(* IEC 61131-3 sources: Caravan/Archiv/12-04-19/Stations/MachineControl/MachineControl/Class/LseEasy (part 2) *)

  if(input < 0) then
    input := 0;
    result := ACCESS_DENIED;
  elsif(input > 100) then
    input := 100;
    result := ACCESS_DENIED;
  else
	  result := input;
  end_if;

  ComPort.SendBacklightDim(input$usint);
	BacklightDim := input;

END_FUNCTION

FUNCTION LseEasy::GetBacklightDim
	VAR_OUTPUT
		retcode 	: USINT;
	END_VAR

  retcode := ComPort.GetBacklightInfo();
  if(retcode <> 0xFF) then
    BacklightDim := retcode and 0x7F;
  end_if;

END_FUNCTION

FUNCTION GLOBAL LseEasy::UpdateScreenshot
	VAR_INPUT
		pscrshot 	: ^void;
	END_VAR

  if(ComPort.SaveScreenshot("C:\hmi35.bmp", pscrshot) = true) then
    OutMessage("SCREENSHOT ...Ready (C:\hmi35.bmp)");
  else
    OutMessage("ERROR: Can't save Screenshot (C:\hmi35.bmp)");
  end_if;

  if(StateSvr = TGetScreenShot) then
    StateSvr := TRun;
  end_if;

END_FUNCTION

FUNCTION VIRTUAL GLOBAL LseEasy::UpdateValue35
	VAR_INPUT
		varno 	: UINT;
		value 	: DINT;
	END_VAR

  if(HmiPrjCrc = Hmi35PrjCrc) then // check crc of project with crc of hmi

    if(varno = VARNO_IRCODE) then
      UpdateIrCode(value$udint);
    end_if;

    HmiVarList.UpdateValue(varno, value);
  end_if;

END_FUNCTION

FUNCTION VIRTUAL GLOBAL LseEasy::UpdateString35
	VAR_INPUT
		varno 	: UINT;
		pstr 	: ^void;
		chrsize 	: UDINT;
	END_VAR

  if(HmiPrjCrc = Hmi35PrjCrc) then // check crc of project with crc of hmi
    HmiVarList.UpdateString(varno, pstr, chrsize);
  end_if;

END_FUNCTION

FUNCTION VIRTUAL GLOBAL LseEasy::UpdateTemperature35
	VAR_INPUT
		value 	: DINT;
	END_VAR

  ActTemperature := value;

END_FUNCTION

FUNCTION GLOBAL LseEasy::UpdateActScreen
	VAR_INPUT
		scrno 	: DINT;
	END_VAR

  ActScreen := scrno;

END_FUNCTION

FUNCTION GLOBAL LseEasy::UpdateInUse

  LastUsage := ops.tAbsolute;

END_FUNCTION

FUNCTION VIRTUAL GLOBAL LseEasy::ActLanguage::Write
	VAR_INPUT
		input (EAX) 	: UDINT;
	END_VAR
	VAR_OUTPUT
		result (EAX) 	: UDINT;
	END_VAR

  if(input <> ActLanguage) then
    if(HmiTextList.GetLanguageIndex(input) <> 16#FFFFFFFF) then
	    ActLanguage := input;
      if(StateSvr = TRun) then
        StateSvr := TStart;
      end_if;
    end_if;
  end_if;

	result := ActLanguage;

END_FUNCTION

FUNCTION GLOBAL LseEasy::SendNewBootLoader
	VAR_OUTPUT
		retcode 	: bool;
	END_VAR

  retcode := SendUpdateToHmi(GetBootLoaderUpdate());

END_FUNCTION

FUNCTION GLOBAL LseEasy::SendNewFirmware
	VAR_OUTPUT
		retcode 	: bool;
	END_VAR

  retcode := SendUpdateToHmi(GetFirmwareUpdate());

END_FUNCTION

FUNCTION LseEasy::SendUpdateToHmi
	VAR_INPUT
		dpne 	: ^CHAR;
	END_VAR
	VAR_OUTPUT
		retcode 	: BOOL;
	END_VAR
  VAR
  	length : udint;
    pbin : ^void;
    tmp : array[0..300] of char;
  END_VAR

  retcode := false;
  pbin    := NIL;

  ComPort.SendBacklightOnOff(1); // turn on backlight

  StringLib.StrCpy(#tmp, 1, "FIRMWARE-UPDATE: Start...[", 1);
  StringLib.StrCat(#tmp, 1, dpne, 1);
  StringLib.StrCat(#tmp, 1, "]", 1);
  OutMessage(#tmp[0]);

  if(File.FOpen(dpne, 'r') = true) then
    length$dint := File.FLength();
    if(length$dint > 0) then
      if(File.FMemory(#pbin, length + 4) = true) then
        if(File.FRead(pbin+4, length) = true) then
          pbin$^udint^ := CRC32_Buffer(pbin+4, length);
          retcode := ComPort.SendNewFirmware(pbin, length+4);
          if(retcode = false) then
            StringLib.StrCpy(#tmp[0], sizeof(char), "ERROR: can't upload ", sizeof(char));
            StringLib.StrCat(#tmp[0], sizeof(char), dpne, sizeof(char));
            OutMessage(#tmp[0]);
          end_if;
        end_if;
        File.FMemory(#pbin, 0);
      end_if;
    end_if;
  else
    StringLib.StrCpy(#tmp[0], sizeof(char), "ERROR: can't open ", sizeof(char));
    StringLib.StrCat(#tmp[0], sizeof(char), dpne, sizeof(char));
    OutMessage(#tmp[0]);
  end_if;

  File.FClose();

  if(retcode = true) then
    OutMessage("FIRMWARE-UPDATE: ...Ready");
  end_if;

END_FUNCTION

FUNCTION GLOBAL LseEasy::SendTrend
	VAR_INPUT
		id 	: UDINT;
		pdata 	: ^USINT;
		length 	: UDINT;
	END_VAR

  ComPort.SendTrendValue(id, pdata, length);

END_FUNCTION

FUNCTION GLOBAL LseEasy::SendPixMap
	VAR_INPUT
		pdata 	: ^void;
		width 	: USINT;
		height 	: USINT;
		padding 	: USINT;
	END_VAR
	VAR_OUTPUT
		retcode 	: BOOL;
	END_VAR
  VAR
  	size : udint;
  END_VAR

  retcode := false;
  size    := ((width * height) + 7) / 8;
  size    += 5; // headerdaten

  // [] ..... command
  // [] ..... version = 1
  // [] ..... width
  // [] ..... height
  // [] ..... padding
  // [ ...... bitdata

  if(size <= sizeof(TmpData)) then
    TmpData[0] := ComCMD_UPDATEPIXMAP;
    TmpData[1] := 1;
    TmpData[2] := width;
    TmpData[3] := height;
    TmpData[4] := padding;
    MemCpy3(#TmpData[5], pdata, size-5);
    retcode := ComPort.SendData(#TmpData[0], size);
  end_if;

END_FUNCTION

FUNCTION GLOBAL LseEasy::OutMessage
	VAR_INPUT
		txt 	: ^CHAR;
	END_VAR
  VAR
  	tmp : array[0..300] of char;
  END_VAR

  tmp[0] := '[';
  tmp[1] := 'N';
  tmp[2] := 'o';
  tmp[3] := 'd';
  tmp[4] := 'e';
  tmp[5] := ' ';
  StringLib.DintToStr(#tmp[6], to_int(ComPort.GetNode()), 16#0800, 1);
  StringLib.StrCat(#tmp[6], 1, "] ", 1);
  StringLib.StrCat(#tmp[6], 1, txt, 1);
  TRACE(#tmp[0]);

END_FUNCTION

FUNCTION LseEasy::OutMessageValue
	VAR_INPUT
		txt 	: ^CHAR;
    value : udint;
	END_VAR
  VAR
  	msg : array[0..128] of char;
  END_VAR

  StringLib.StrCpy(#msg[0], 1, txt, 1);
  StringLib.DintToStr(#msg[StringLib.StrLen(#msg[0], 1)], to_dint(value), 0x800, 1);
  OutMessage(#msg[0]);

END_FUNCTION

FUNCTION GLOBAL LseEasy::UpdateAll
	VAR_INPUT
		act_hmi_crc 	: UDINT;
	END_VAR

  Hmi35PrjCrc   := act_hmi_crc;
  NeedUpdateAll += 1;

END_FUNCTION

FUNCTION LseEasy::CheckCrc
VAR
	crc : udint;
END_VAR

  crc := ComPort.GetFileCrc(0);
  if(crc = 16#FFFFFFFF) then
    // there is no valid project in hmi
    StateSvr := TStart; // restart
  elsif(crc <> 0) then
    CantGetCrc := 0;
    if(crc = HmiPrjCrc) then
      // same project detected in hmi
      UpdateAll(crc); // force update of all data
      StateSvr := TRun;
    else
      // different project detected in hmi
      StateSvr := TStart; // restart
    end_if;
  else

    SleepNext(StateSvr, 100); // sleep 100ms

    CantGetCrc += 1;
    if(CantGetCrc > 100) then
      CantGetCrc := 0;
      ErrorStateSvr(true);
    end_if;
  end_if;

END_FUNCTION

FUNCTION GLOBAL LseEasy::UpdateAliveSignal35

  AliveTix35     := ops.tAbsolute;
  HmiOnline      := 1;
  AliveTix35Cntr += 1;

END_FUNCTION

FUNCTION GLOBAL LseEasy::UpdateBacklight35
	VAR_INPUT
		state 	: DINT;
	END_VAR

//  if(state and 0x80) then
//    BacklightOnOff := 1;
//  else
//    BacklightOnOff := 0;
//  end_if;

  BacklightDim := state and 0x7F;

END_FUNCTION

FUNCTION LseEasy::CheckProjectCrc
	VAR_INPUT
		ptr 	: ^void;
		hmiver 	: UDINT;
		chkold 	: bool;
	END_VAR
	VAR_OUTPUT
		retcode 	: BOOL;
	END_VAR
  VAR
  	pprj : ^_BOX_PROJECTLIST;
  	phlp : ^_BOX_PROJECTLIST_ENTRY;
    no, index : udint;
		pbox	: ^_BIGBOX_HEADER;
    upload : bool;
  END_VAR

  upload     := true;
  retcode    := false;
  pbox$^void := ptr;

  if(ComPort.GetFileCrc(0) = pbox^.crc32) then
    retcode := true;
    upload  := false;
    if((chkold = true) & (hmiver < 127)) then
      // einzelne crc's im hmi überprüfen
      // erst ab hmi-version 1.27 werden die crc's mit GetFileCrc(0) direkt im hmi überprüft
      pprj$^void := pbox;
      no         := pprj^.no;
      phlp       := #pprj^.data[0];
      index      := 0;

      while(no) do
        no    -= 1;
        pbox$^void := HmiProject35.GetBox(index);

        if(ComPort.GetFileCrc(phlp^.filename) <> pbox^.crc32) then
          retcode := false;
          no      := 0;
        end_if;

        phlp  += sizeof(_BOX_PROJECTLIST_ENTRY);
        index += 1;
      end_while;
    end_if;
  end_if;

  if(IsProjectUpLoadNecessary(upload) = true) then
    retcode := false;
  end_if;

END_FUNCTION

FUNCTION LseEasy::SendProject
	VAR_INPUT
		ptr 	: ^void;
	END_VAR
	VAR_OUTPUT
		retcode 	: BOOL;
	END_VAR
  VAR
  	pprj : ^_BOX_PROJECTLIST;
  	phlp : ^_BOX_PROJECTLIST_ENTRY;
    no, index, tix, nox, sizeram, sizeflash : udint;
    pbox : ^_BIGBOX_HEADER;
    upload : bool;
  END_VAR

  retcode := false;
  upload  := false;

  tix := ops.tAbsolute;

    if(ComPort.SendReset() = true) then

      HmiSwVersion := ComPort.GetSwVersion();
      HmiHwVersion := ComPort.GetHwVersion();

      GetBacklightDim();

      pbox$^void := ptr;
      retcode    := true;

      // nur wenn projektcrc unterschiedlich
      if(CheckProjectCrc(ptr, HmiSwVersion, false) = false) then

        if(ComPort.GetHardwareData(nil, #sizeram, #sizeflash) = true) then
          sizeflash := sizeflash - (24 + 512*16); // flashhader + fatgrösse abziehen
          if((HmiProject35.TotalByteSize > sizeflash) | (HmiProject35.TotalFileNo > 256)) then
            OutMessage("ERROR: Size of LSE-Project is too big");
            OutMessageValue("...PrjSize[byte] = ", HmiProject35.TotalByteSize);
            OutMessageValue("...MaxSize[byte] = ", sizeflash);
            SetErrorSvr(ErrSizeLseProject);
            retcode := false;
          end_if;
        end_if;

        if(retcode = true) then

          // clear flash
          if(ComPort.SendFormatFlash() = true) then

            OutMessage("HMI-UPDATE: Start...");

            // send projectentries
            pprj$^void := ptr;
            no         := pprj^.no;
            phlp       := #pprj^.data[0];
            index      := 0;
//            totalsize  := 0;

            while(no) do
              ComPort.ShowProgressBar(to_usint((index * 100) / pprj^.no));

              no    -= 1;
              pbox$^void := HmiProject35.GetBox(index);

              if(ComPort.SendFile(phlp^.filename, pbox^.size, pbox) = false) then
                OutMessageValue("ERROR: Upload ProjectEntry of Bytesize = ", pbox^.size);
                retcode := false;
                no      := 0;
              end_if;
//              totalsize += HmiProject35.AlignU32(pbox^.size);
              phlp  += sizeof(_BOX_PROJECTLIST_ENTRY);
              index += 1;
            end_while;

            if(retcode = true) then
              // send projektlist
              ComPort.ShowProgressBar(100);
              pbox$^void := ptr;
              retcode    := ComPort.SendFile(0, pbox^.size, pbox);
//              totalsize  += HmiProject35.AlignU32(pbox^.size);

              if(retcode = true) then
                HmiMapFile.Create(GetPrjPath(), pbox^.crc32);
                OutMessageValue("HMI-UPDATE: ...Ready, TotalSize[byte] = ", HmiProject35.TotalByteSize); //totalsize);
                // vorsicht: projekt ist jetzt im hmi-ram, noch nicht auf flash
                retcode := ComPort.Ping(); // send ping to ensure alive-hmi and update alivetrigger
              end_if;
              upload := true;
            end_if;

          else
            retcode := false;
          end_if;
        end_if;
      end_if;

      if(retcode = true) then
        UpdateAll(HmiPrjCrc); // force updateall
        nox := ops.tAbsolute;
        repeat
          if(ComPort.SendRun() = true) then
            exit;
          end_if;
        until((ops.tAbsolute - nox) > 1000) end_repeat;

        if(upload = true) then
          // after performing projectupload, sleep a while to ensure flash of whole project-data in hmi
          nox := ops.tAbsolute;
          while((ops.tAbsolute - nox) < 1000) do
          end_while;
          ComPort.Ping(); // send ping to keep hmi happy
        end_if;

        OutMessageValue("HMI-RUN: UpdateTime[ms] = ", ops.tAbsolute - tix);
      else
        OutMessage("ERROR: Upload HMI-Project");
        SetErrorSvr(ErrUploadHmiProject);
        ComPort.SendChkTraceView(); // display message on hmi
      end_if;
    end_if;

END_FUNCTION

FUNCTION LseEasy::Run

  // alivesignal
  if((ops.tabsolute - AliveTix) > 1003) then
    AliveTix := ops.tabsolute;
    ComPort.SendAliveTrigger(); // send alive trigger to hmi
  end_if;

  // onlinewatchdog
  if((ops.tabsolute - AliveTix35) > 4000) then
    HmiOnline := 0; // offline
    if(TempInterval <> 0) then
      ActTemperature$UDINT := 0x80000010; // fühlerbruch
    end_if;
  end_if;

  if(HmiOnline) then

    if(HmiPrjCrc = Hmi35PrjCrc) then // check crc of project with crc of hmi

      if(NeedUpdateAll) then
        NeedUpdateAll := 0;
        GetBacklightDim();
        HmiVarList.RefreshAll();
        HmiStateBit35.RefreshAll();
        HmiReady();
      end_if;

      HmiRun();

      if((ops.tabsolute - RefreshTix) > 6) then
        RefreshTix := ops.tAbsolute;
        HmiVarList.RefreshRun();
        HmiStateBit35.RefreshRun();
      end_if;

      if(TrendVal0 <> -1) then
        TrendVal0 := UpdateTrendVal(0, TrendVal0);
      end_if;

      if(TrendVal1 <> -1) then
        TrendVal1 := UpdateTrendVal(1, TrendVal1);
      end_if;

      if(PixMap <> -1) then
        PixMap := UpdatePixMap(PixMap);
      end_if;

    else
      // just in this moment we're back online with hmi
      SleepNext(TChkCrc, 1000); // wait a while and afterwards check project
    end_if;
  else
    Hmi35PrjCrc := 0; // destroy hmicrc
    CantGetCrc  := 0;
  end_if;

  if(CallScreen <> -1) then
    if(CallScreen = -2) then
      OutMessage("SCREENSHOT: Start...");
      if(ComPort.GetScreenShot() = false) then
        OutMessage("ERROR: Screenshot not done");
      else
        StateSvr := TGetScreenShot;
      end_if;
    else
      ComPort.SendGotoScreen(CallScreen);
    end_if;
    CallScreen := -1;
  end_if;

END_FUNCTION

FUNCTION VIRTUAL GLOBAL LseEasy::Background
	VAR_INPUT
		EAX 	: UDINT;
	END_VAR
	VAR_OUTPUT
		state (EAX) 	: UDINT;
	END_VAR

	state := READY;

  case StateSvr of
    TStart :
      AutoFirmwareUpdate := AutoFirmwareUpdate.Read();
      if(ComPort.Ping() = true) then // ask for hmi
        if(LoadFile() = true) then
          if(Create() = true) then
            StateSvr := TUpload;
          end_if;
        end_if;

        if(StateSvr <> TUpload) then
          ErrorStateSvr(false);
        else
          if(AutoFirmwareUpdate <> 0) then
            if(AutoFwUpdateDisabled = false) then
              AutoFwUpdateDisabled := true; // no further auto-update of firmware possible
              StateSvr := TCheckUpdateBootloader;
            end_if;
          end_if;
        end_if;
      else
        OutMessage("ERROR: Can't communicate with HMI");
        SetErrorSvr(ErrHmiCommunication);
        ErrorStateSvr(true);
      end_if;

    TCheckUpdateBootLoader :
      StateSvr := CheckUpdate(GetBootloaderUpdate(), TCheckUpdateFirmware, TCheckUpdateFirmware, 15000);

    TCheckUpdateFirmware :
      StateSvr := CheckUpdate(GetFirmwareUpdate(), TStart, TUpLoad, 17000);

    TUpLoad :
      if(UpLoadProject() = true) then
        HmiProject35.Free();
        ProjectBox := NIL;
        StateSvr := TRun;
      end_if;

    TGetScreenShot :
      Run();

    TRun :
      Run();

    TFirmwareUpdate :
      if(SendNewFirmware() = true) then
        SleepNext(TRun, 10000);
      else
        ErrorStateSvr(false);
      end_if;

    TBootLoaderUpdate :
      if(SendNewBootLoader() = true) then
        SleepNext(TRun, 10000);
      else
        ErrorStateSvr(false);
      end_if;

    TChkCrc :
      CheckCrc();

    TSleep :
      if((ops.tAbsolute - SleepStart) >= SleepDuration) then
        StateSvr := StateNext;
      end_if;

    TReboot :
      ComPort.SendReboot();
      SleepNext(TStart, 3000);

    TError :
      if(TryToRestart = true) then
        if(AliveTix35Cntr <> AliveTix35CntrOld) then
          // try to restart after hmi sent alivesignal
          StateSvr     := TStart;
          TryToRestart := false;
        end_if;
      end_if;

  end_case;

  ComPort.Run();

END_FUNCTION

FUNCTION VIRTUAL GLOBAL LseEasy::StateSvr::Write
	VAR_INPUT
		input (EAX) 	: LseEasy::TStateSvr;
	END_VAR
	VAR_OUTPUT
		result (EAX) 	: LseEasy::TStateSvr;
	END_VAR

  if(input = TGetScreenShot) then
    result$udint := ACCESS_DENIED;
    if(StateSvr = TRun) then
      CallScreen := -2;
	    result     := StateSvr;
    end_if;
  else
	  StateSvr := input;
	  result := StateSvr;
  end_if;

END_FUNCTION

FUNCTION VIRTUAL GLOBAL LseEasy::HmiAccess
	VAR_INPUT
		level 	: UDINT;
	END_VAR
	VAR_OUTPUT
		retcode 	: BOOL;
	END_VAR

  retcode := true;
  if(level > AccessLevel) then
    retcode := false;
  end_if;

END_FUNCTION

FUNCTION GLOBAL LseEasy::SoftReset

  StateSvr := TStart;

END_FUNCTION

FUNCTION GLOBAL LseEasy::SoftResetAll
  VAR
  	nox : udint;
    pth : ^LseEasy;
  END_VAR

  pth := InstancePtr[0];
  nox := InstanceCnt;
  while(nox) do
    pth^.SoftReset();
    nox -= 1;
    pth += sizeof(InstancePtr[0]);
  end_while;

END_FUNCTION

FUNCTION VIRTUAL GLOBAL LseEasy::ClassSvr::NewInst
	VAR_INPUT
		pPara 	: ^CmdStruct;
		pResult 	: ^Results;
	END_VAR
	VAR_OUTPUT
		ret_code 	: IprStates;
	END_VAR

	ret_code := READY;

	case pPara^.uiCmd of

		0 : // start download on the fly
        pResult^.aData[0]$UDINT := 16#46544F44; // DOTF-id
        pResult^.uiLng          := 6; // success

		1 : // end download on the fly
        pResult^.aData[0]$UDINT := 16#46544F44; // DOTF-id
        pResult^.uiLng          := 6; // success
        SoftResetAll();
  end_case;

END_FUNCTION

#pragma warning (disable : 73)
FUNCTION VIRTUAL GLOBAL LseEasy::UserCall
	VAR_INPUT
		fktno 	: UDINT;
		para 	: DINT;
	END_VAR

END_FUNCTION
#pragma warning (default : 73)

#pragma warning (disable : 73)
FUNCTION VIRTUAL GLOBAL LseEasy::HmiVariableExtention
	VAR_INPUT
		varname 	: ^CHAR;
	END_VAR
	VAR_OUTPUT
		retcode 	: UDINT;
	END_VAR

  retcode := 16#FFFFFFFF;

//  if(StringLib.StrCmp(varname, sizeof(char), "Dummy.Server7", sizeof(char)) = 0) then
//    retcode := VARNO_TEST_NUM1;
//  end_if;

END_FUNCTION
#pragma warning (default : 73)

FUNCTION LseEasy::GetMapCrc
	VAR_OUTPUT
		retcode 	: UDINT;
	END_VAR

  retcode := HmiVarList.GetMapCrc();
  retcode := (retcode rol 1) xor HmiStateBit35.GetMapCrc();

END_FUNCTION

FUNCTION VIRTUAL LseEasy::IsProjectUpLoadNecessary
	VAR_INPUT
		preselect 	: BOOL;
	END_VAR
	VAR_OUTPUT
		retcode 	: BOOL;
	END_VAR

//  if(GetmapCrc() <> oldmapcrc) then
    // unconditional upload necessary, otherwise weak functionality of hmi
//  end_if;

  retcode := preselect;

END_FUNCTION

FUNCTION VIRTUAL GLOBAL LseEasy::UpdatePixMap
	VAR_INPUT
		value 	: DINT;
	END_VAR
	VAR_OUTPUT
		retcode 	: DINT;
	END_VAR

  retcode := value;
  if(SendPixMap(#value, 32, 1, 0) = true) then
    retcode := -1;
  end_if;

END_FUNCTION

FUNCTION VIRTUAL GLOBAL LseEasy::UpdateTrendVal
	VAR_INPUT
    id : UDINT;
		value 	: DINT;
	END_VAR
	VAR_OUTPUT
		retcode 	: DINT;
	END_VAR

  retcode := value;
  if(ComPort.SendTrendValue(id, #(value$usint), 1) = true) then
    retcode := -1;
  end_if;

END_FUNCTION

FUNCTION LseEasy::Recalculate_MulDiv
	VAR_INPUT
		einheit 	: UDINT;
		posdezpt 	: DINT;
	END_VAR
	VAR_OUTPUT
		retcode 	: DINT;
	END_VAR
  var
    dekade : dint;
  end_var

  retcode := 1;
  dekade  := 0;

  case(einheit) of
    1000000000 : dekade := 9;
    100000000  : dekade := 8;
    10000000   : dekade := 7;
    1000000    : dekade := 6;
    100000     : dekade := 5;
    10000      : dekade := 4;
    1000       : dekade := 3;
    100        : dekade := 2;
    10         : dekade := 1;
  end_case;

  case(dekade - posdezpt) of
    9 : retcode := 1000000000;
    8 : retcode :=  100000000;
    7 : retcode :=   10000000;
    6 : retcode :=    1000000;
    5 : retcode :=     100000;
    4 : retcode :=      10000;
    3 : retcode :=       1000;
    2 : retcode :=        100;
    1 : retcode :=         10;
  end_case;

END_FUNCTION

FUNCTION LseEasy::Recalculate_Calc
	VAR_INPUT
		rval 	: real;
    rmul  : real;
		rdiv 	: real;
		direction 	: bool;
	END_VAR
	VAR_OUTPUT
		retcode 	: DINT;
	END_VAR

  if(direction = true) then
    rval := (rval * rmul) / rdiv;
  else
    rval := (rval * rdiv) / rmul;
  end_if;

  retcode := to_dint(rval);

//  if(rval < 0) then
//    retcode := to_dint(rval - 0.5);
//  else
//    retcode := to_dint(rval + 0.5);
//  end_if;

END_FUNCTION

FUNCTION VIRTUAL LseEasy::Recalculate_Stroke2mm
  VAR_INPUT
    value : DINT;
    dezpoint : DINT;
    direction : BOOL;
  END_VAR
  VAR_OUTPUT
    retcode : DINT;
  END_VAR
  VAR
  	rdiv : real;
  END_VAR

  rdiv    := Recalculate_MulDiv(1mm, dezpoint);
  retcode := Recalculate_Calc(value, 1.0, rdiv, direction);

END_FUNCTION

FUNCTION VIRTUAL LseEasy::Recalculate_Stroke2inch
  VAR_INPUT
    value : DINT;
    dezpoint : DINT;
    direction : BOOL;
  END_VAR
  VAR_OUTPUT
    retcode : DINT;
  END_VAR
  VAR
  	rdiv : real;
  END_VAR

  rdiv    := Recalculate_MulDiv(1mm, dezpoint);
  retcode := Recalculate_Calc(value, 1.0, rdiv * 25.4, direction);

END_FUNCTION

FUNCTION VIRTUAL LseEasy::Recalculate_Temp2Celsius
  VAR_INPUT
    value : DINT;
    dezpoint : DINT;
    direction : BOOL;
  END_VAR
  VAR_OUTPUT
    retcode : DINT;
  END_VAR
  VAR
  	rdiv : real;
  END_VAR

  rdiv    := Recalculate_MulDiv(10, dezpoint);
  retcode := Recalculate_Calc(value, 1.0, rdiv, direction);

END_FUNCTION

FUNCTION VIRTUAL LseEasy::Recalculate_Temp2Fahrenheit
  VAR_INPUT
    value : DINT;
    dezpoint : DINT;
    direction : BOOL;
  END_VAR
  VAR_OUTPUT
    retcode : DINT;
  END_VAR

  if(direction = true) then
    if(value < 0) then
      retcode := ((value * 18 - 5) / 10) + 320;
    else
      retcode := ((value * 18 + 5) / 10) + 320;
    end_if;

    if(dezpoint = 0) then
      if(value < 0) then
        retcode := (retcode - 5) / 10;
      else
        retcode := (retcode + 5) / 10;
      end_if;
    elsif(dezpoint = 2) then
      retcode := retcode * 10;
    end_if;
  else
    if(dezpoint = 0) then
      value := value * 10;
    elsif(dezpoint = 2) then
      if(value < 0) then
        value := (value - 5) / 10;
      else
        value := (value + 5) / 10;
      end_if;
    end_if;

    if(value < 0) then
      retcode := (((value - 320) * 10) - 9) / 18;
    else
      retcode := (((value - 320) * 10) + 9) / 18;
    end_if;

  end_if;

END_FUNCTION

FUNCTION VIRTUAL LseEasy::Recalculate_Weight2Kilogram
  VAR_INPUT
    value : DINT;
    dezpoint : DINT;
    direction : BOOL;
  END_VAR
  VAR_OUTPUT
    retcode : DINT;
  END_VAR
  VAR
  	rdiv : real;
  END_VAR

  rdiv    := Recalculate_MulDiv(10000, dezpoint);
  retcode := Recalculate_Calc(value, 1.0, rdiv, direction);

END_FUNCTION

FUNCTION VIRTUAL LseEasy::Recalculate_Weight2Pound
  VAR_INPUT
    value : DINT;
    dezpoint : DINT;
    direction : BOOL;
  END_VAR
  VAR_OUTPUT
    retcode : DINT;
  END_VAR
  VAR
  	rdiv : real;
  END_VAR

  rdiv    := Recalculate_MulDiv(10000, dezpoint);
  retcode := Recalculate_Calc(value, 2.204622, rdiv, direction);

END_FUNCTION

FUNCTION VIRTUAL LseEasy::Recalculate_Pressure2Bar
  VAR_INPUT
    value : DINT;
    dezpoint : DINT;
    direction : BOOL;
  END_VAR
  VAR_OUTPUT
    retcode : DINT;
  END_VAR
  VAR
  	rdiv : real;
  END_VAR

  rdiv    := Recalculate_MulDiv(1bar, dezpoint);
  retcode := Recalculate_Calc(value, 1.0, rdiv, direction);

END_FUNCTION

FUNCTION VIRTUAL LseEasy::Recalculate_Pressure2Psi
  VAR_INPUT
    value : DINT;
    dezpoint : DINT;
    direction : BOOL;
  END_VAR
  VAR_OUTPUT
    retcode : DINT;
  END_VAR
  VAR
  	rdiv : real;
  END_VAR

  rdiv    := Recalculate_MulDiv(1bar, dezpoint);
  retcode := Recalculate_Calc(value, 14.50376808, rdiv, direction);

END_FUNCTION

FUNCTION VIRTUAL LseEasy::Recalculate_Time2Second
  VAR_INPUT
    value : DINT;
    dezpoint : DINT;
    direction : BOOL;
  END_VAR
  VAR_OUTPUT
    retcode : DINT;
  END_VAR

  retcode := Recalculate_MulDiv(1sec, dezpoint);

  if(direction = true) then
    if(value < 0) then
      retcode := (value - (retcode / 2)) / retcode;
    else
      retcode := (value + (retcode / 2)) / retcode;
    end_if;
  else
    retcode := value * retcode;
  end_if;

END_FUNCTION

FUNCTION VIRTUAL LseEasy::Recalculate_Time2Minute
  VAR_INPUT
    value : DINT;
    dezpoint : DINT;
    direction : BOOL;
  END_VAR
  VAR_OUTPUT
    retcode : DINT;
  END_VAR

  if(direction = true) then
    if(value < 0) then
      retcode := Recalculate_Time2Second((value - 30) / 60, dezpoint, true);
    else
      retcode := Recalculate_Time2Second((value + 30) / 60, dezpoint, true);
    end_if;
  else
    retcode := Recalculate_Time2Second(value * 60, dezpoint, false);
  end_if;

END_FUNCTION

FUNCTION VIRTUAL LseEasy::Recalculate_Time2Hour
  VAR_INPUT
    value : DINT;
    dezpoint : DINT;
    direction : BOOL;
  END_VAR
  VAR_OUTPUT
    retcode : DINT;
  END_VAR

  if(direction = true) then
    if(value < 0) then
      retcode := Recalculate_Time2Minute((value - 30) / 60, dezpoint, true);
    else
      retcode := Recalculate_Time2Minute((value + 30) / 60, dezpoint, true);
    end_if;
  else
    retcode := Recalculate_Time2Minute(value * 60, dezpoint, false);
  end_if;

END_FUNCTION

FUNCTION VIRTUAL LseEasy::Recalculate_Force2KN
  VAR_INPUT
    value : DINT;
    dezpoint : DINT;
    direction : BOOL;
  END_VAR
  VAR_OUTPUT
    retcode : DINT;
  END_VAR
  VAR
  	rdiv : real;
  END_VAR

  rdiv    := Recalculate_MulDiv(1kn, dezpoint);
  retcode := Recalculate_Calc(value, 1.0, rdiv, direction);

END_FUNCTION

FUNCTION VIRTUAL GLOBAL LseEasy::Recalculate
	VAR_INPUT
		value 	: DINT;
		formula 	: UDINT;
		dezpoint 	: DINT;
		direction 	: BOOL;
	END_VAR
	VAR_OUTPUT
		retcode 	: DINT;
	END_VAR

  retcode := value;

  case formula of
    3  : retcode := Recalculate_Stroke2mm(value, dezpoint, direction);
    4  : retcode := Recalculate_Stroke2inch(value, dezpoint, direction);
    5  : retcode := Recalculate_Temp2Celsius(value, dezpoint, direction);
    6  : retcode := Recalculate_Temp2Fahrenheit(value, dezpoint, direction);
    7  : retcode := Recalculate_Weight2Kilogram(value, dezpoint, direction);
    8  : retcode := Recalculate_Weight2Pound(value, dezpoint, direction);
    9  : retcode := Recalculate_Pressure2Bar(value, dezpoint, direction);
    10 : retcode := Recalculate_Pressure2Psi(value, dezpoint, direction);
    11 : retcode := Recalculate_Time2Second(value, dezpoint, direction);
    12 : retcode := Recalculate_Time2Minute(value, dezpoint, direction);
    13 : retcode := Recalculate_Time2Hour(value, dezpoint, direction);
    14 : retcode := Recalculate_Force2KN(value, dezpoint, direction);
  end_case;

END_FUNCTION

FUNCTION GLOBAL LseEasy::SoftResetIn
	VAR_INPUT
		milliseconds 	: UDINT;
	END_VAR

  SleepNext(TStart, milliseconds);

END_FUNCTION

#pragma warning (disable : 73)
FUNCTION VIRTUAL LseEasy::UpdateIrCode
	VAR_INPUT
		code 	: UDINT;
	END_VAR

END_FUNCTION
#pragma warning (default : 73)

FUNCTION VIRTUAL GLOBAL LseEasy::CheckUpdate
	VAR_INPUT
		dpne 	: ^CHAR;
		nextstep 	: TStateSvr;
		defaultstep 	: TStateSvr;
		sleep 	: UDINT;
	END_VAR
	VAR_OUTPUT
		retcode 	: TStateSvr;
	END_VAR

  retcode := defaultstep;

  if(File.FOpen(dpne, 'r') = true) then // is updatefile present
    File.FClose();
    if(SendUpdateToHmi(dpne) = true) then
      if(AutoFirmwareUpdate = 1) then
        File.FDelete(dpne); // delete file
      end_if;
      retcode := SleepNext(nextstep, sleep);
    end_if;
  end_if;

END_FUNCTION

FUNCTION GLOBAL  LseEasy::GetLseProjectNotice
	VAR_OUTPUT
		retcode 	: ^char;
	END_VAR

  retcode := HmiSetUpList.GetLseProjectNotice();

END_FUNCTION
